// Balise pilotée par le séquenceur auquel elle est rattachée (docs/02 § 8, docs/03 § 8.1)
INTERFACE I_Beacon

METHOD SetPattern
VAR_INPUT
    nPattern : UINT;             // bits de F_BeaconBits
    bBuzzer : BOOL;
END_VAR
END_METHOD

END_INTERFACE

(* stored: Version 1.1.0.1, ProductVersion 3.1.4024.12
   Itf I_Beacon: Id {70016109-5c95-5508-85c7-55da30e90c25}
   Method SetPattern: Id {341c0480-23ab-58fb-97e1-f88919af11b7} *)
